FUNCTION_BLOCK stop (* Basic Function Block Type *)
  (* Standard: 61499-2 *)
  (* Version 0.0, 10/21/2026, lizar, Schneider Electric, Template *)
  PACKAGE Main;
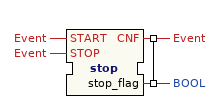
  EVENT_INPUT
    START; (* Initialization Request *)
    STOP; (* Normal Execution Request *)
  END_EVENT
  EVENT_OUTPUT
    CNF WITH stop_flag; (* Execution Confirmation *)
  END_EVENT
  VAR_OUTPUT
    stop_flag : BOOL; (* Output event qualifier *)
  END_VAR
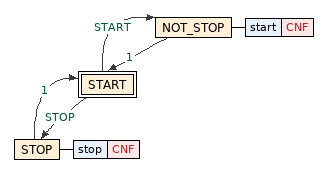
  EC_STATES
    START; (* Initial State *)
    NOT_STOP : start -> CNF; (* Initialization *)
    STOP : stop -> CNF; (* Normal execution *)
  END_STATES
  EC_TRANSITIONS
    START TO NOT_STOP := START;
    NOT_STOP TO START := 1;
    START TO STOP := STOP;
    STOP TO START := 1;
  END_TRANSITIONS
  ALGORITHM stop IN ST: (* Initialization algorithm *)
;
stop_flag:=TRUE;
  END_ALGORITHM
  ALGORITHM start IN ST:
;
stop_flag:=FALSE;
  END_ALGORITHM
END_FUNCTION_BLOCK
